FUNCTION_BLOCK FB_Prototype
VAR
	nCount	: INT;
END_VAR

nCount := nCount + UnknownSymbol; // not built: the folder is excluded from the build

END_FUNCTION_BLOCK

(* stored: Version 1.1.0.1
   POU FB_Prototype: Id {6bc0fb70-9147-4b8d-9dc2-36f739b84163}, SpecialFunc None *)
